FUNCTION_BLOCK PhaseEmergencyStart (* Basic Function Block Type *)
  (* Standard: 61499-2 *)
  (* Version 0.1, 28/10/2026, Schneider Electric, 0.1: entrada Mode; no EmergencyOFF a fase rodando recebe parada se o modo ainda for 3. *)
  PACKAGE SE.Nereda;
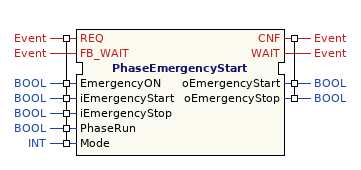
  EVENT_INPUT
    REQ WITH iEmergencyStart, iEmergencyStop, PhaseRun, EmergencyON, Mode; (* Normal Execution Request *)
    FB_WAIT;
  END_EVENT
  EVENT_OUTPUT
    CNF WITH oEmergencyStart, oEmergencyStop; (* Execution Confirmation *)
    WAIT;
  END_EVENT
  VAR_INPUT
    EmergencyON : BOOL;
    iEmergencyStart : BOOL; (* Input event qualifier *)
    iEmergencyStop : BOOL;
    PhaseRun : BOOL;
    Mode : INT; (* Modo atual (3 = emergencia); lido no REQ *)
  END_VAR
  VAR_OUTPUT
    oEmergencyStart : BOOL; (* Output event qualifier *)
    oEmergencyStop : BOOL;
  END_VAR
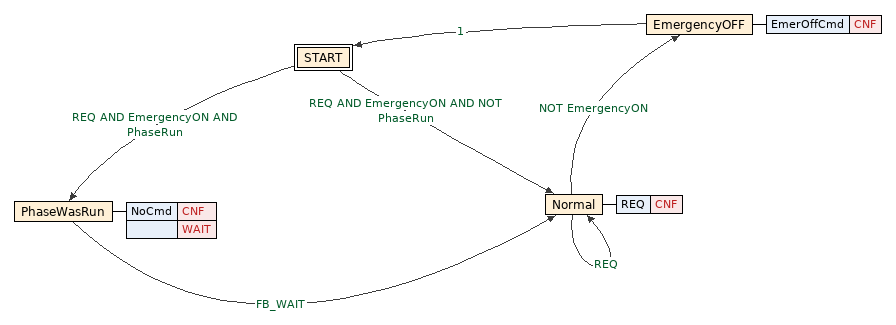
  EC_STATES
    START; (* Initial State *)
    PhaseWasRun : NoCmd -> CNF, -> WAIT;
    Normal : REQ -> CNF;
    EmergencyOFF : EmerOffCmd -> CNF;
  END_STATES
  EC_TRANSITIONS
    Normal TO EmergencyOFF := NOT EmergencyON;
    START TO PhaseWasRun := REQ AND EmergencyON AND PhaseRun;
    START TO Normal := REQ AND EmergencyON AND NOT PhaseRun;
    PhaseWasRun TO Normal := FB_WAIT;
    Normal TO Normal := REQ;
    EmergencyOFF TO START := 1;
  END_TRANSITIONS
  ALGORITHM REQ IN ST: (* Normally executed algorithm *)
;
oEmergencyStart := iEmergencyStart;
oEmergencyStop := iEmergencyStop;
  END_ALGORITHM
  ALGORITHM EmerOffCmd IN ST: (* Emergencia desligada para esta fase *)
;
(* Reator saiu da emergencia com o modo ainda em 3 (indisponivel / forcado indisponivel):
   a fase que estava rodando para. Se o modo ja saiu de 3, nao manda nada (Nereda / operador assume). *)
oEmergencyStart := FALSE;
oEmergencyStop := PhaseRun AND (Mode = 3);
  END_ALGORITHM
  ALGORITHM NoCmd IN ST:
;
oEmergencyStart := FALSE;
oEmergencyStop := FALSE;
  END_ALGORITHM
END_FUNCTION_BLOCK
